{attribute 'qualified_only'}
// Interface contract
INTERFACE I_Device EXTENDS I_Base

METHOD ReadValue : BOOL
VAR_INPUT
    channel : INT;
END_VAR
END_METHOD

PROPERTY Enabled : BOOL
GET
END_GET
SET
END_SET
END_PROPERTY

METHOD Reset
END_METHOD

END_INTERFACE

(* stored: Version 1.1.0.1
   Itf I_Device: Id {b7f34f64-9ec4-43e3-92ca-41e3431d02a1} *)
